// TIA Portal V17 export
FUNCTION_BLOCK "BeltRun"   // FB, LAD
// Runs the belt.
   VAR_INPUT
      StartButton : Bool;   // Start button
      StopButton : Bool;   // Stop button
   END_VAR
   VAR_OUTPUT
      BeltMotor : Bool;   // Belt motor
   END_VAR
BEGIN

REGION Network 1: Run the belt
   // Start turns the belt on when stop is off.
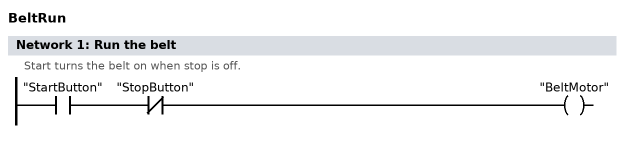
   RUNG wire#powerrail
      Contact( "StartButton" )
      I_Contact( "StopButton" )
      Coil( "BeltMotor" )
   END_RUNG
   // the same network as SCL:
   "BeltMotor" := "StartButton" AND NOT "StopButton";
END_REGION
END_FUNCTION_BLOCK

FUNCTION "ScaleLevel" : Void   // FC, FBD
   VAR_INPUT
      Level : Real;   // Tank level
      Offset : Real;   // Speed offset
   END_VAR
   VAR_OUTPUT
      Result : Real;   // Scaled result
   END_VAR
BEGIN

REGION Network 1: Add the offset
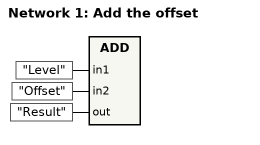
   <??.?> := "Level" + "Offset" + "Result";
END_REGION
END_FUNCTION

ORGANIZATION_BLOCK "FillPump"   // OB, SCL
   VAR
      Level : Real;   // Tank level
      Pump : Bool;   // Fill pump
   END_VAR
BEGIN
// Fill when the level is low
   IF "Level" < 10 THEN "Pump" := TRUE;
END_ORGANIZATION_BLOCK

FUNCTION_BLOCK "FillSequence"   // FB, GRAPH
BEGIN
// Fill then discharge
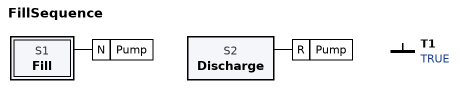
   // sequencer 1
   INITIAL_STEP Fill:   // S1
              N    Pump
   END_STEP
   STEP Discharge:   // S2
              R    Pump
   END_STEP
   TRANSITION "" FROM ? TO ?   // T1
      := TRUE;
   END_TRANSITION
END_FUNCTION_BLOCK
